(* CODESYS project system.library
   DefaultNamespace: KOSTAL.TC3.Core.System
   DocFormat: reStructuredText
   Description: Contains basic definitions for an OOP construction.
   Author: Frank Dümpelmann
   Title: KOSTAL.TC3.Core.System
   Version: 2019.0.0.0
   Company: KOSTAL GmbH & Co.KG
   Placeholder: KOSTAL.TC3.Core.System

Project tree, tasks and I/O mapping:
  Interface/
    interface I_Interface
  Project Information/
    function F_GetCompany [ST]
    function F_GetTitle [ST]
    function F_GetVersion [ST]
  Version/
    global variables Global_Version
*)

// Version/Global_Version
{attribute 'TcGenerated'}
{attribute 'no-analysis'}
{attribute 'linkalways'}
// This function has been automatically generated from the project information.
VAR_GLOBAL CONSTANT
	{attribute 'const_non_replaced'}
	stLibVersion_KOSTAL_TC3_Core_System : ST_LibVersion := (iMajor := 2019, iMinor := 0, iBuild := 0, iRevision := 0, nFlags := 0, sVersion := '2019.0.0.0');
END_VAR

// Interface/I_Interface
(*
	Base Interface for all basic interfaces in KOSTAL.TC3. Interfaces
*)
INTERFACE I_Interface EXTENDS __SYSTEM.IQueryInterface

END_INTERFACE

// Project Information/F_GetCompany
// This function has been automatically generated from the project information.
{attribute 'signature_flag' := '1073741824'}
{attribute 'TcGenerated'}
{attribute 'no-analysis'}
FUNCTION F_GetCompany : WSTRING
VAR_INPUT
	
END_VAR

F_GetCompany := "KOSTAL GmbH & Co.KG";

END_FUNCTION

// Project Information/F_GetTitle
// This function has been automatically generated from the project information.
{attribute 'signature_flag' := '1073741824'}
{attribute 'TcGenerated'}
{attribute 'no-analysis'}
FUNCTION F_GetTitle : WSTRING
VAR_INPUT
	
END_VAR

F_GetTitle := "KOSTAL.TC3.Core.System";

END_FUNCTION

// Project Information/F_GetVersion
// This function has been automatically generated from the project information.
{attribute 'signature_flag' := '1073741824'}
{attribute 'TcGenerated'}
{attribute 'no-analysis'}
FUNCTION F_GetVersion : ST_LibVersion
VAR_INPUT
	
END_VAR

F_GetVersion.iMajor := 2019;
F_GetVersion.iMinor := 0;
F_GetVersion.iBuild := 0;
F_GetVersion.iRevision := 0;
F_GetVersion.sVersion := '2019.0.0.0';
F_GetVersion.nFlags := 0;

END_FUNCTION
